Fanuc KAREL source: KA00123.KL

PROGRAM KA00123
%NOLOCKGROUP
VAR
  SRC: ARRAY[2] OF BYTE
  DST: BOOLEAN
BEGIN
  SRC[1] = 2
  DST = SRC[1]
END KA00123
